// TIA Portal V19 export
FUNCTION_BLOCK "DRIVE_RPM"   // FB45, LAD
{ S7_Optimized_Access := 'TRUE' }
// stored: MemoryReserve 100, SetENOAutomatically false
   VAR_INPUT
      RAW_MIN : Array[1..20] of Int;
      RAW_MAX : Array[1..20] of Int;
      SCALE_MIN : Array[1..20] of Real;
      SCALE_MAX : Array[1..20] of Real;
      INPUT : Array[1..20] of Int;
   END_VAR
   VAR_OUTPUT
      FAULT : Array[1..20] of Bool;
      SCALE_OUT : Array[1..20] of Real;
      STATUS : Array[1..20] of Int;
   END_VAR
   VAR
      AI : Array[1..20] of "SCALING";
      MAX_VALUE { S7_SetPoint := 'True'} : Array[1..20] of Int;
      I : Int;
   END_VAR
BEGIN

REGION Network 1 (SCL)

   FOR #I := 1 TO 20 DO
       IF #INPUT[#I] < -100 OR #INPUT[#I] > 28648 THEN
           #FAULT[#I] := 1;
       ELSE
           #FAULT[#I] := 0;
       END_IF;
       IF NOT #FAULT[#I] THEN
           #AI[#I](RAW_MIN := #RAW_MIN[#I],
                   RAW_MAX := #RAW_MAX[#I],
                   INPUT := #INPUT[#I],
                   SCALE_MIN := #SCALE_MIN[#I],
                   SCALE_MAX := #SCALE_MAX[#I],
                   SCALE_OUT => #SCALE_OUT[#I]);
       ELSE
           #SCALE_OUT[#I] := 0.0;

       END_IF;


       IF #SCALE_OUT[#I]>3 THEN
           #STATUS[#I] := 1;
       ELSE
           #STATUS[#I] := 2;

       END_IF;

       ;
   END_FOR;
END_REGION
END_FUNCTION_BLOCK
